# EPICS substitutions: iocs/motor/acsmotion-ioc/db/AcsMotionAuxIO.substitutions
# C's iocAcsMotion AcsMotionAuxIO.substitutions, P and PORT (the
# AcsMotionAuxIOConfig port) from st.cmd.

file "$(ACSMOTION_IOC)/db/SPiiPlusAuxLi.db"
{
pattern
{C,     R,   CHAN, SCAN}
# MP4U
{mp4u:, li0, 0,    2}
{mp4u:, li1, 1,    2}
{mp4u:, li2, 2,    2}
{mp4u:, li3, 3,    2}
}

file "$(ACSMOTION_IOC)/db/SPiiPlusAuxLo.db"
{
pattern
{C,     R,   CHAN, SCAN}
# MP4U
{mp4u:, lo0, 0,    2}
{mp4u:, lo1, 1,    2}
{mp4u:, lo2, 2,    2}
{mp4u:, lo3, 3,    2}
}

file "$(ACSMOTION_IOC)/db/SPiiPlusAuxBi.db"
{
pattern
{C,     R,      CHAN, MASK,    SCAN}
# MP4U
{mp4u:, bi0:17, 0,    0x10000, 2}
{mp4u:, bi0:18, 0,    0x20000, 2}
{mp4u:, bi0:19, 0,    0x40000, 2}
{mp4u:, bi0:20, 0,    0x80000, 2}
{mp4u:, bi1:17, 1,    0x10000, 2}
{mp4u:, bi1:18, 1,    0x20000, 2}
{mp4u:, bi1:19, 1,    0x40000, 2}
{mp4u:, bi1:20, 1,    0x80000, 2}
{mp4u:, bi2:17, 2,    0x10000, 2}
{mp4u:, bi2:18, 2,    0x20000, 2}
{mp4u:, bi2:19, 2,    0x40000, 2}
{mp4u:, bi2:20, 2,    0x80000, 2}
{mp4u:, bi3:17, 3,    0x10000, 2}
{mp4u:, bi3:18, 3,    0x20000, 2}
{mp4u:, bi3:19, 3,    0x40000, 2}
{mp4u:, bi3:20, 3,    0x80000, 2}
}

file "$(ACSMOTION_IOC)/db/SPiiPlusAuxBo.db"
{
pattern
{C,     R,     CHAN, MASK,  SCAN}
# MP4U
{mp4u:, bo0:8, 0,    0x100, 2}
{mp4u:, bo0:9, 0,    0x200, 2}
{mp4u:, bo1:8, 1,    0x100, 2}
{mp4u:, bo1:9, 1,    0x200, 2}
{mp4u:, bo2:8, 2,    0x100, 2}
{mp4u:, bo2:9, 2,    0x200, 2}
{mp4u:, bo3:8, 3,    0x100, 2}
{mp4u:, bo3:9, 3,    0x200, 2}
}

file "$(ACSMOTION_IOC)/db/SPiiPlusAuxAo.db"
{
pattern
{C,     R,    CHAN, SCAN, DRVL, DRVH, LOPR, HOPR, PREC}
# MP4U
{mp4u:, ao0,  0,    2,    -10,  10,   -10,  10,   3}
{mp4u:, ao1,  1,    2,    -10,  10,   -10,  10,   3}
{mp4u:, ao2,  2,    2,    -10,  10,   -10,  10,   3}
{mp4u:, ao3,  3,    2,    -10,  10,   -10,  10,   3}
{mp4u:, ao4,  4,    2,    -10,  10,   -10,  10,   3}
{mp4u:, ao5,  5,    2,    -10,  10,   -10,  10,   3}
{mp4u:, ao6,  6,    2,    -10,  10,   -10,  10,   3}
{mp4u:, ao7,  7,    2,    -10,  10,   -10,  10,   3}
{mp4u:, ao8,  8,    2,    -10,  10,   -10,  10,   3}
{mp4u:, ao9,  9,    2,    -10,  10,   -10,  10,   3}
{mp4u:, ao10, 10,   2,    -10,  10,   -10,  10,   3}
{mp4u:, ao11, 11,   2,    -10,  10,   -10,  10,   3}
{mp4u:, ao12, 12,   2,    -10,  10,   -10,  10,   3}
{mp4u:, ao13, 13,   2,    -10,  10,   -10,  10,   3}
{mp4u:, ao14, 14,   2,    -10,  10,   -10,  10,   3}
{mp4u:, ao15, 15,   2,    -10,  10,   -10,  10,   3}
# IOMps-EA0004V0
{mp4u:, ao16, 16,   2,    -10,  10,   -10,  10,   3}
{mp4u:, ao17, 17,   2,    -10,  10,   -10,  10,   3}
{mp4u:, ao18, 18,   2,    -10,  10,   -10,  10,   3}
{mp4u:, ao19, 19,   2,    -10,  10,   -10,  10,   3}
}

file "$(ACSMOTION_IOC)/db/SPiiPlusAuxAi.db"
{
pattern
{C,     R,    CHAN, SCAN, LOPR, HOPR, PREC}
# MP4U
{mp4u:, ai0,  0,    2,    -10,  10,   3}
{mp4u:, ai1,  1,    2,    -10,  10,   3}
{mp4u:, ai2,  2,    2,    -10,  10,   3}
{mp4u:, ai3,  3,    2,    -10,  10,   3}
{mp4u:, ai4,  4,    2,    -10,  10,   3}
{mp4u:, ai5,  5,    2,    -10,  10,   3}
{mp4u:, ai6,  6,    2,    -10,  10,   3}
{mp4u:, ai7,  7,    2,    -10,  10,   3}
{mp4u:, ai8,  8,    2,    -10,  10,   3}
{mp4u:, ai9,  9,    2,    -10,  10,   3}
{mp4u:, ai10, 10,   2,    -10,  10,   3}
{mp4u:, ai11, 11,   2,    -10,  10,   3}
{mp4u:, ai12, 12,   2,    -10,  10,   3}
{mp4u:, ai13, 13,   2,    -10,  10,   3}
{mp4u:, ai14, 14,   2,    -10,  10,   3}
{mp4u:, ai15, 15,   2,    -10,  10,   3}
}
